// Parameters of FB TON and FB TOF.
TYPE
ST_SafeTimerParameters :
STRUCT
    MakeContact : BOOL;
    DelayTime : TIME;
END_STRUCT
END_TYPE

(* stored: Version 1.1.0.1
   DUT ST_SafeTimerParameters: Id {6ccc2540-9b4a-56c2-8b2e-2d65f34748b1} *)
